(* Schneider Machine Expert - Basic project m221 plc, file version 2.9.0.0 *)
(* ProjectInformations: Name=New project *)

HARDWARE
  Cpu 0: TM221CE24R
  EthernetConfiguration: NetworkName=M221, IpAllocationMode=FixedAddress, IpAddress=192.168.1.113, SubnetMask=255.255.255.0
  SerialLineConfiguration: Baud=Baud19200, Parity=ParityEven, DataBits=DataBits8, StopBits=StopBits1, PhysicalMedium=PhysicalMediumRs485, TransmissionMode=TransmissionModeModbusRtu, SlaveId=1, Addressing=SlaveAddressing
  MastTask: UsePeriodScanMode=false, PeriodScan=100
  FastTask: Period=255
  CpuBehavior: StartingMode=StartAsPreviousState, AutoSaveRamOnEeprom=true, WatchdogPeriod=250

SYMBOLS  (address, symbol, comment, settings)
  %M0       START_1
  %M1       STOP1
  %M2       START_2
  %M3       STOP_2
  %M4       RUN1
  %M5       RUN2
  %I0.0     REMOTE1
  %I0.1     REMOTE2
  %I0.2     ESTOP
  %Q0.0     VSD1
  %Q0.1     VSD2

POU New POU
  (* SectionNumber=1 *)

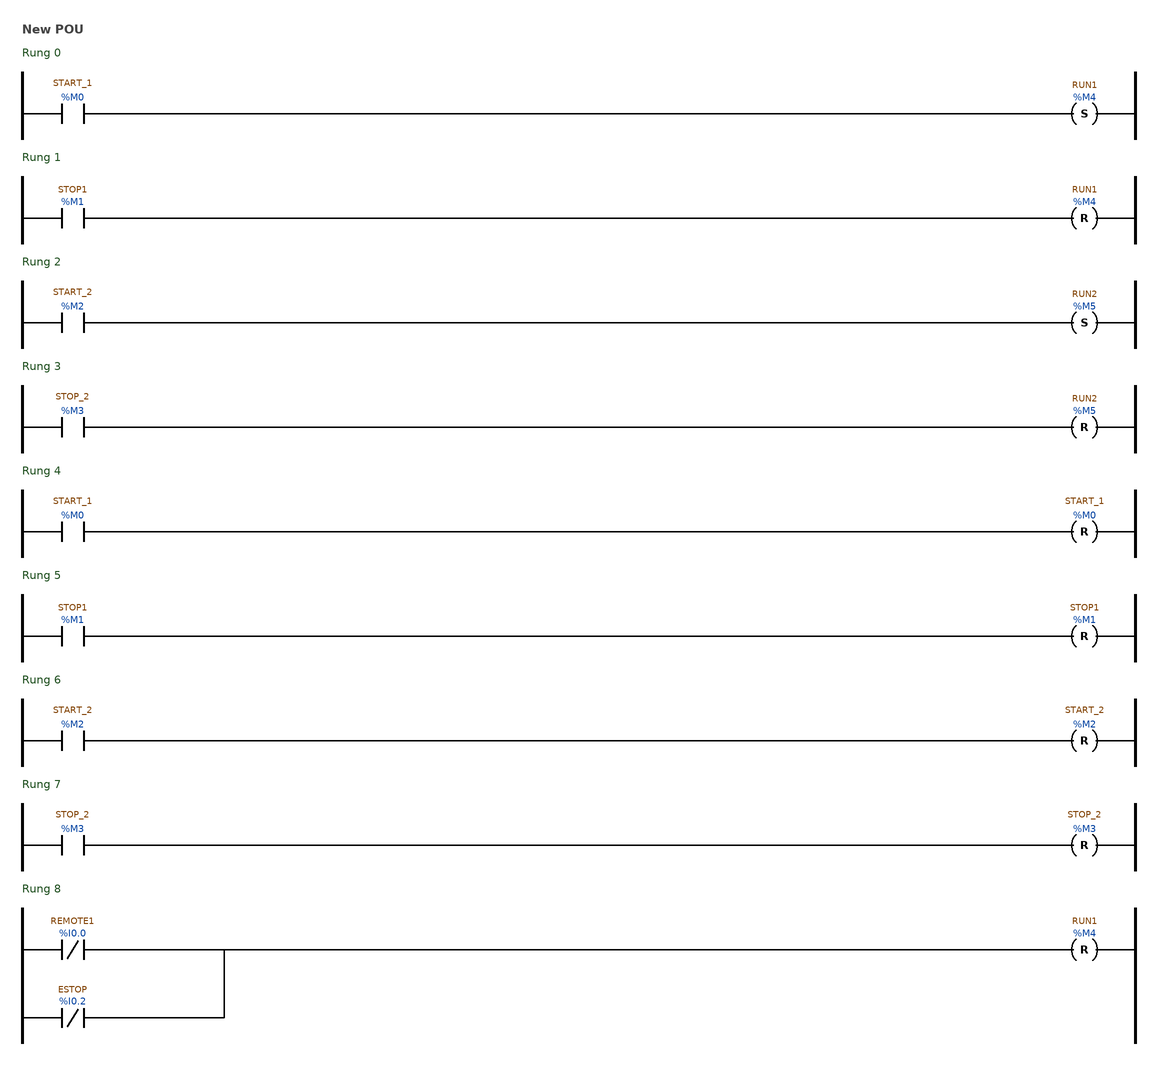

// Rung 0
  LD %M0                  (* START_1 *)
  S %M4                   (* RUN1 *)
  // as ST:
  //   IF START_1 THEN RUN1 := TRUE; END_IF;

// Rung 1
  LD %M1                  (* STOP1 *)
  R %M4                   (* RUN1 *)
  // as ST:
  //   IF STOP1 THEN RUN1 := FALSE; END_IF;

// Rung 2
  LD %M2                  (* START_2 *)
  S %M5                   (* RUN2 *)
  // as ST:
  //   IF START_2 THEN RUN2 := TRUE; END_IF;

// Rung 3
  LD %M3                  (* STOP_2 *)
  R %M5                   (* RUN2 *)
  // as ST:
  //   IF STOP_2 THEN RUN2 := FALSE; END_IF;

// Rung 4
  LD %M0                  (* START_1 *)
  R %M0                   (* START_1 *)
  // as ST:
  //   IF START_1 THEN START_1 := FALSE; END_IF;

// Rung 5
  LD %M1                  (* STOP1 *)
  R %M1                   (* STOP1 *)
  // as ST:
  //   IF STOP1 THEN STOP1 := FALSE; END_IF;

// Rung 6
  LD %M2                  (* START_2 *)
  R %M2                   (* START_2 *)
  // as ST:
  //   IF START_2 THEN START_2 := FALSE; END_IF;

// Rung 7
  LD %M3                  (* STOP_2 *)
  R %M3                   (* STOP_2 *)
  // as ST:
  //   IF STOP_2 THEN STOP_2 := FALSE; END_IF;

// Rung 8
  LDN %I0.0               (* REMOTE1 *)
  ORN %I0.2               (* ESTOP *)
  R %M4                   (* RUN1 *)
  // as ST:
  //   IF NOT REMOTE1 OR NOT ESTOP THEN RUN1 := FALSE; END_IF;

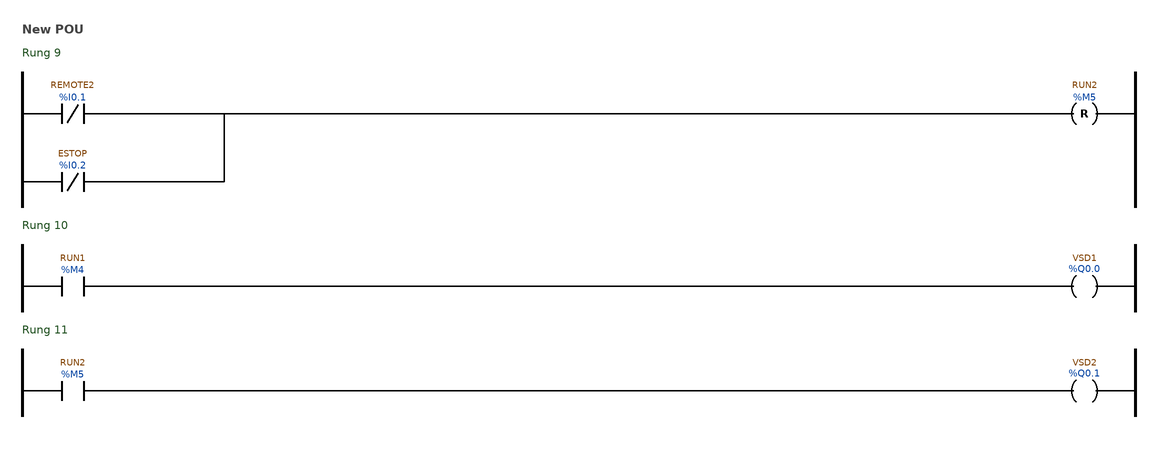

// Rung 9
  LDN %I0.1               (* REMOTE2 *)
  ORN %I0.2               (* ESTOP *)
  R %M5                   (* RUN2 *)
  // as ST:
  //   IF NOT REMOTE2 OR NOT ESTOP THEN RUN2 := FALSE; END_IF;

// Rung 10
  LD %M4                  (* RUN1 *)
  ST %Q0.0                (* VSD1 *)
  // as ST:
  //   VSD1 := RUN1;

// Rung 11
  LD %M5                  (* RUN2 *)
  ST %Q0.1                (* VSD2 *)
  // as ST:
  //   VSD2 := RUN2;
